(*
SPDX-FileCopyrightText: © 2026 Oleksandr Tiutyk <trofimich@gmail.com>
SPDX-License-Identifier: MIT
License: https://opensource.org/license/mit
*)

(*!
<summary>Combines one or more child workflow conditions using a logical AND or OR operator.</summary>
<description>
Requires at least one child condition to be considered Configured. Short-circuits evaluation on the first
decisive child result.
</description>
*)

{attribute 'no_explicit_call' := 'do not call this function block directly'}
{attribute 'enable_dynamic_creation'}
FUNCTION_BLOCK CompositeCondition EXTENDS Condition IMPLEMENTS ICompositeCondition, TOF_Core.IConfigurationSerializable
VAR_STAT
	{attribute 'hide'}
	_ClassName : STRING := __POUNAME();
END_VAR
VAR
	{attribute 'OPC.UA.DA' := '0'}
	_LogicalOperator : LOGICAL_OPERATOR;

	{attribute 'OPC.UA.DA' := '0'}
	_Children : TOF_Collections.List<0>(valueValidator := 0);
END_VAR

(*!
<summary>Appends a child condition and assigns this composite as its ParentCondition.</summary>
<description>
Rejects null references, self/ancestor cycles and conditions already attached elsewhere.
The child must be unattached, including to this parent; duplicate slots are rejected before insertion.
The parent chain and owning workflow must be PASSIVE_READY. Fixed workflow association is validated.
Storage allocation precedes parent callbacks; callback exceptions may leave a partial configuration.
Child references remain borrowed and must outlive the tree. No implicit detach or ownership transfer occurs.
</description>
<param name="condition">Child condition to append.</param>
*)
METHOD AddChildCondition
VAR_INPUT
	condition : ICondition;
END_VAR
VAR
	childParent : IWorkflowElement;
END_VAR
IF condition = 0 THEN
	TOF_Core.Exceptions.ThrowArgumentNotSpecified(
		sourceNamespaceName := NamespaceName,
		sourceClassName := ClassName,
		sourcePOUName := __POUNAME(),
		sourcePosition := __POSITION(),
		argumentName := 'condition'
	);
END_IF

Workflows.ValidateElementAttachment(parent := THIS^, child := condition);

childParent := condition.Parent;

IF childParent <> 0 THEN
	WorkflowExceptions.ThrowWorkflowAttachment(
		sourceNamespaceName := NamespaceName,
		sourceClassName := ClassName,
		sourcePOUName := __POUNAME(),
		sourcePosition := __POSITION(),
		message := "Child element already occupies a parent slot"
	);
END_IF

_Children.AppendGeneric(
	value := TOF_Core.GenericValueFactory.FromParts(
		genericTypeClass := TOF_Core.GENERIC_TYPE_CLASS.OBJECT,
		address := condition.SelfAddress,
		size := condition.SelfSize,
		memoryManagementBehavior := TOF_Core.GENERIC_MEMORY_MANAGEMENT_BEHAVIOR.STORE_ORIGINAL_REFERENCE_AND_NOT_OWNS_MEMORY
	)
);

condition.ParentCondition := THIS^;
END_METHOD

(*!
<summary>Borrows the initialized class name used in diagnostics.</summary>
<description>
Returns initialized metadata storage without allocation. Callers must not modify the returned string.
Derived function blocks must use distinct initialized static storage when overriding this metadata.
</description>
*)
{attribute 'monitoring' := 'call'}
PROPERTY ClassName : REFERENCE TO STRING
GET
ClassName REF= _ClassName;
END_GET
END_PROPERTY

(*!
<summary>Returns TRUE when at least one child condition has been added.</summary>
*)
{attribute 'monitoring' := 'call'}
PROPERTY Configured : BOOL
GET
Configured := _Children.Length > TOF_Core.SignedInt32.ZERO;
END_GET
END_PROPERTY

(*!
<summary>Gets or sets the logical operator (AND_ or OR_) used to combine child conditions.</summary>
*)
PROPERTY LogicalOperator : LOGICAL_OPERATOR
GET
LogicalOperator := _LogicalOperator;
END_GET
SET
_LogicalOperator := LogicalOperator;
END_SET
END_PROPERTY

(*!
<summary>Borrows the compiler-initialized library namespace.</summary>
<description>
Borrows storage from the live internal namespace provider. Reacquire references after application
reinitialization or relocation. Treat the reference as read-only; no ownership or synchronization is provided.
</description>
*)
{attribute 'monitoring' := 'call'}
PROPERTY NamespaceName : REFERENCE TO STRING
GET
NamespaceName REF= CurrentNamespace.Name;
END_GET
END_PROPERTY

(*!
<summary>Evaluates child conditions in order and short-circuits according to LogicalOperator.</summary>
<param name="activity">Activity context for evaluation.</param>
*)
METHOD PROTECTED OnEvaluate : BOOL
VAR_INPUT
	activity : IActivity;
END_VAR
VAR
	formattedExceptionMessage : TOF_Core.ERROR_MESSAGE;


	i : DINT;
	
	childCondition : ICondition;
END_VAR
IF NOT Configured THEN
	formattedExceptionMessage := TOF_Core.WideStrings.Concat255("Condition '", Name, "' is not configured");

	WorkflowExceptions.ThrowWorkflowConfiguration(
		sourceNamespaceName := NamespaceName,
		sourceClassName := ClassName,
		sourcePOUName := __POUNAME(),
		sourcePosition := __POSITION(),
		message := formattedExceptionMessage
	);
END_IF

IF _LogicalOperator = LOGICAL_OPERATOR.AND_ THEN
	OnEvaluate := TRUE;
END_IF

FOR i := 0 TO _Children.Length - 1 DO
	IF NOT __QUERYINTERFACE(_Children.Get(index := i).AsObject(), childCondition) THEN
		formattedExceptionMessage := TOF_Core.WideStrings.Concat255("Condition #", TO_WSTRING(i), " is null");

		WorkflowExceptions.ThrowWorkflowConfiguration(
			sourceNamespaceName := NamespaceName,
			sourceClassName := ClassName,
			sourcePOUName := __POUNAME(),
			sourcePosition := __POSITION(),
			message := formattedExceptionMessage
		);
	END_IF

	IF NOT childCondition.Configured THEN
		formattedExceptionMessage := TOF_Core.WideStrings.Concat255(
			"Condition '",
			childCondition.Name,
			"' is not configured"
		);

		WorkflowExceptions.ThrowWorkflowConfiguration(
			sourceNamespaceName := NamespaceName,
			sourceClassName := ClassName,
			sourcePOUName := __POUNAME(),
			sourcePosition := __POSITION(),
			message := formattedExceptionMessage
		);
	END_IF

	IF childCondition.Evaluate(activity := activity) THEN
		IF _LogicalOperator = LOGICAL_OPERATOR.OR_ THEN
			OnEvaluate := TRUE;
			RETURN;
		END_IF
	ELSE
		IF _LogicalOperator = LOGICAL_OPERATOR.AND_ THEN
			OnEvaluate := FALSE;
			RETURN;
		END_IF
	END_IF
END_FOR
END_METHOD

(*!
<summary>Reports the size of this concrete function block instance in bytes.</summary>
<description>
Reports the instance layout rather than dynamic allocations owned by its fields. A derived function block
with a different layout must override this property; the value does not grant disposal rights.
</description>
*)
{attribute 'monitoring' := 'call'}
PROPERTY SelfSize : ULINT
GET
SelfSize := XSIZEOF(THIS^);
END_GET
END_PROPERTY

(*!
<summary>Writes the configuration fields for this object.</summary>
<description>Borrows the writer for this call. A failure invalidates the current output document.</description>
*)
METHOD Serialize
VAR_INPUT
	writer : TOF_Core.IConfigurationWriter;
END_VAR
VAR
	operatorText : STRING;
	i : DINT;
END_VAR
Workflows.WriteConfigurationHeader(writer := writer, source := THIS^, displayName := Name, scope := THIS^);
operatorText := Workflows.FormatLogicalOperator(logicalOperator := _LogicalOperator);
writer.WriteValue(
	name := 'operator',
	valueType := TOF_Core.CONFIGURATION_VALUE_TYPE.TYPE_STRING,
	data := ADR(operatorText),
	size := SIZEOF(operatorText)
);
writer.BeginArray(name := 'children');

FOR i := 0 TO _Children.Length - 1 DO
	Workflows.WriteConfigurationObject(writer := writer, name := '', source := _Children.Get(index := i).AsObject());
END_FOR

writer.EndArray();
END_METHOD

(*!
<summary>Restores this fresh instance from its configuration object.</summary>
<description>
The reader, document node and deserialization context are borrowed for this call.
On failure discard the partial instance.
</description>
<param name="reader">Active configuration reader.</param>
<param name="node">Object node to read fields from.</param>
<param name="context">Active configuration deserialization context providing workflow reconstruction services.</param>
*)
METHOD Deserialize
VAR_INPUT
	reader : TOF_Core.IConfigurationReader;
	node : TOF_Core.CONFIGURATION_NODE;
	context : TOF_Core.IConfigurationDeserializationContext;
END_VAR
VAR
	loader : IWorkflowLoader;
	items : TOF_Core.CONFIGURATION_NODE;
	count : DINT;
	i : DINT;
	operatorText : STRING;
END_VAR
loader := WorkflowConfigurationSerializer.ResolveWorkflowLoader(context := context);
Workflows.ReadConfigurationHeader(reader := reader, node := node, target := THIS^, scope := THIS^);

operatorText := Workflows.ReadName(
	reader := reader,
	node := reader.GetField(node := node, name := 'operator')
);
LogicalOperator := Workflows.ParseLogicalOperator(rawOperator := operatorText);

items := reader.GetField(node := node, name := 'children');
count := TO_DINT(reader.GetArraySize(node := items));

FOR i := 0 TO count - 1 DO
	AddChildCondition(
		condition := Workflows.ReadCondition(loader := loader, node := reader.GetItem(node := items, index := TO_UDINT(i)))
	);
END_FOR
END_METHOD

END_FUNCTION_BLOCK

(* stored: Version 1.1.0.1
   POU CompositeCondition: Id {8a55c5b1-693f-4932-9f9a-010c3c539516}, SpecialFunc None
   Folder Overriden methods: Id {92167edf-a171-45ae-b0b4-cbb4363d35a0}
   Method AddChildCondition: Id {a9ba8ac8-dab1-4579-a8c6-f1dcf4f0781e}
   Property ClassName: Id {70333ea1-3549-4d0a-a3ad-521d1db0db74}
   Get Get: Id {a5ccd782-e1de-457e-9e73-065fb67a7a80}
   Property Configured: Id {21dacc3f-ed62-4ab7-8da9-cb67ea9bfcba}
   Get Get: Id {ea5c9fa4-9f95-445e-834b-d8986cf079b5}
   Property LogicalOperator: Id {2e60dc3a-8843-4578-a90f-416536b1cdcb}
   Get Get: Id {24be606b-b29e-4d7a-9059-3d33397fc9bc}
   Set Set: Id {91bb16fb-1705-4e7d-aeac-ee32b7347b30}
   Property NamespaceName: Id {52983f0a-5112-4343-a340-1487d5e77845}
   Get Get: Id {8a11a0fb-561b-4d9a-b1ae-2ae3af60f58b}
   Method OnEvaluate: Id {65421d01-d63f-414e-ae6f-3caad321436b}
   Property SelfSize: Id {0c774fc8-e3e1-46bd-bc7e-7d6910760a9c}
   Get Get: Id {02bdd4c2-e6e9-4e38-a963-e1672ee8a20b}
   Method Serialize: Id {4ae6e667-f885-4f73-a2bf-809bae770cbb}
   Method Deserialize: Id {e594c35e-bafc-4c07-b96d-dc9ce4cf9508} *)
